Fanuc KAREL source: kt00585.KL

-- PROVISIONAL review KL for V1013-1; original PC SHA256 a276833919a1b081c0a67a75b49e65dfa11f25616956c5f822ced15fbe681812
-- Incomplete behavior may be omitted. Consult companion uncertainty JSON. Do not deploy.
PROGRAM KT00585
%NOLOCKGROUP
VAR
  I1 : INTEGER
-- UNRESOLVED_DECL V2 type=000013
-- UNRESOLVED_DECL OUT type=000013
BEGIN
  -- UNRESOLVED_PC offsets 5-16; opcodes 2E,23
  -- UNRESOLVED_PC offsets 21-36; opcodes 2E,22,32,35
  -- UNRESOLVED_PC offsets 41-63; opcodes 21,49,8B,4A
  -- UNRESOLVED_PC offsets 68-72; opcodes 7F
END KT00585
